// Mitsubishi GX Works2 project: 공개1번(FX)   PLC: FX3U/FX3UC

PROGRAM MAIN
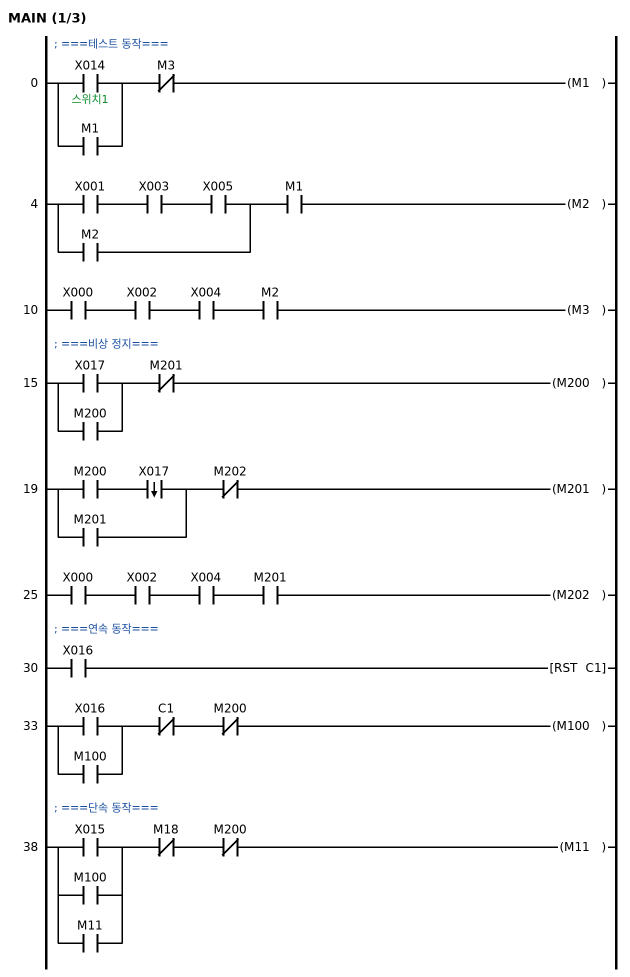
; ===테스트 동작===
0     LD      X014  ; 스위치1
      OR      M1
      ANI     M3
      OUT     M1
4     LD      X001
      AND     X003
      AND     X005
      OR      M2
      AND     M1
      OUT     M2
10    LD      X000
      AND     X002
      AND     X004
      AND     M2
      OUT     M3
; ===비상 정지===
15    LD      X017
      OR      M200
      ANI     M201
      OUT     M200
19    LD      M200
      ANDF    X017
      OR      M201
      ANI     M202
      OUT     M201
25    LD      X000
      AND     X002
      AND     X004
      AND     M201
      OUT     M202
; ===연속 동작===
30    LD      X016
      RST     C1
33    LD      X016
      OR      M100
      ANI     C1
      ANI     M200
      OUT     M100
; ===단속 동작===
38    LD      X015
      OR      M100
      OR      M11
      ANI     M18
      ANI     M200
      OUT     M11
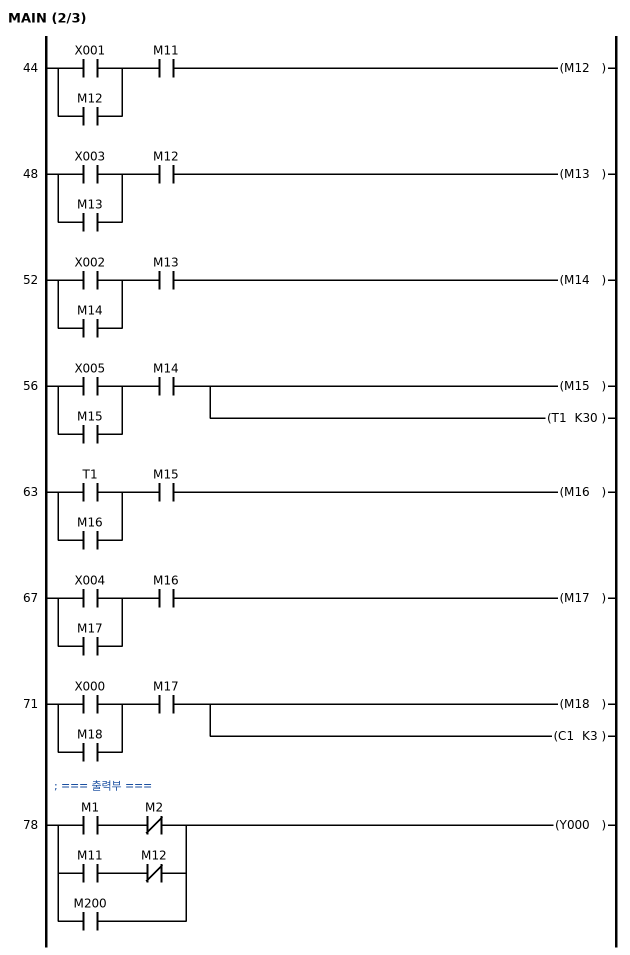
44    LD      X001
      OR      M12
      AND     M11
      OUT     M12
48    LD      X003
      OR      M13
      AND     M12
      OUT     M13
52    LD      X002
      OR      M14
      AND     M13
      OUT     M14
56    LD      X005
      OR      M15
      AND     M14
      OUT     M15
      OUT     T1 K30
63    LD      T1
      OR      M16
      AND     M15
      OUT     M16
67    LD      X004
      OR      M17
      AND     M16
      OUT     M17
71    LD      X000
      OR      M18
      AND     M17
      OUT     M18
      OUT     C1 K3
; === 출력부 ===
78    LD      M1
      ANI     M2
      LD      M11
      ANI     M12
      ORB
      OR      M200
      OUT     Y000
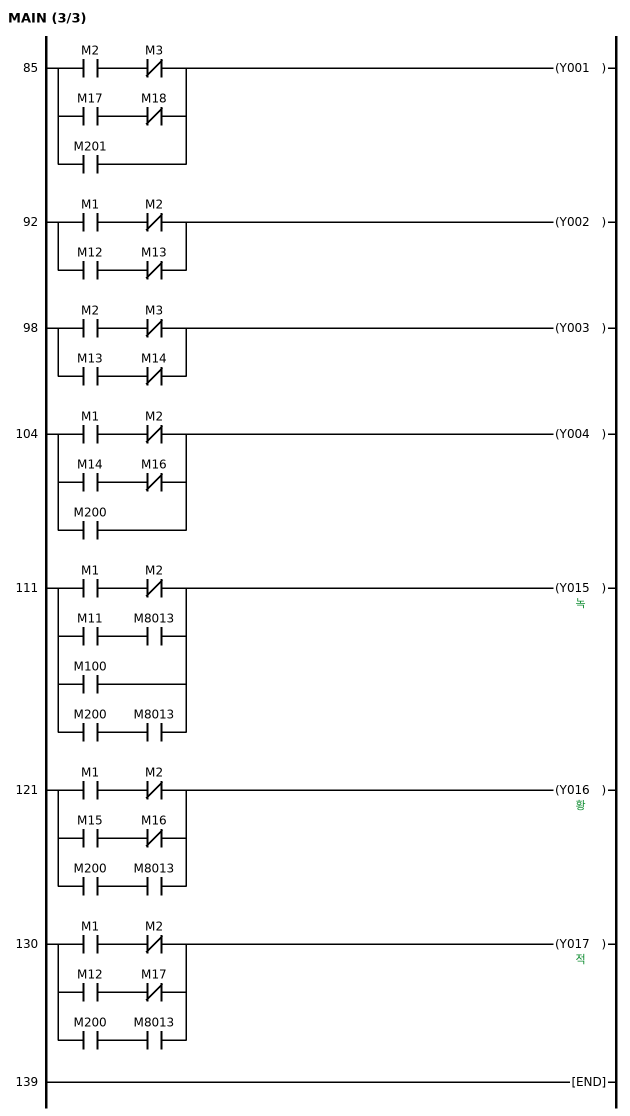
85    LD      M2
      ANI     M3
      LD      M17
      ANI     M18
      ORB
      OR      M201
      OUT     Y001
92    LD      M1
      ANI     M2
      LD      M12
      ANI     M13
      ORB
      OUT     Y002
98    LD      M2
      ANI     M3
      LD      M13
      ANI     M14
      ORB
      OUT     Y003
104   LD      M1
      ANI     M2
      LD      M14
      ANI     M16
      ORB
      OR      M200
      OUT     Y004
111   LD      M1
      ANI     M2
      LD      M11
      AND     M8013
      ORB
      OR      M100
      LD      M200
      AND     M8013
      ORB
      OUT     Y015  ; 녹
121   LD      M1
      ANI     M2
      LD      M15
      ANI     M16
      ORB
      LD      M200
      AND     M8013
      ORB
      OUT     Y016  ; 황
130   LD      M1
      ANI     M2
      LD      M12
      ANI     M17
      ORB
      LD      M200
      AND     M8013
      ORB
      OUT     Y017  ; 적
139   END
END_PROGRAM
